// TIA Portal V20 export
DATA_BLOCK "OP2_DB"   // DB1
// stored: InstanceOfName OP2, InstanceOfType FB
"OP2"
   // VAR
   //    CONTROL_MAN : Struct
   //       B0 : Bool;
   //       B1 : Bool;
   //       B2 : Bool;
   //       B3 : Bool;
   //       B4 : Bool;
   //       B5 : Bool;
   //       B6 : Bool;
   //       B7 : Bool;
   //       B8 : Bool;
   //       B9 : Bool;
   //       odfuk_1 : Bool;
   //       odfuk_2 : Bool;
   //       B12 : Bool;
   //       B13 : Bool;
   //       B14 : Bool;
   //       B15 : Bool;
   //       B16 : Bool;
   //       B17 : Bool;
   //       B18 : Bool;
   //       B19 : Bool;
   //       B20 : Bool;
   //       B21 : Bool;
   //       B22 : Bool;
   //       B23 : Bool;
   //       B24 : Bool;
   //       B25 : Bool;
   //       B26 : Bool;
   //       B27 : Bool;
   //       B28 : Bool;
   //       B29 : Bool;
   //       B30 : Bool;
   //       B31 : Bool;
   //    END_STRUCT;
   //    CONTROL_AUTOMAT : Struct
   //       connect : Bool;
   //       send : Bool;
   //       reciv : Bool;
   //       trcv : Bool;
   //       discon : Bool;
   //       B5 : Bool;
   //       B6 : Bool;
   //       B7 : Bool;
   //       B8 : Bool;
   //       B9 : Bool;
   //       B10 : Bool;
   //       B11 : Bool;
   //       B12 : Bool;
   //       B13 : Bool;
   //       B14 : Bool;
   //       B15 : Bool;
   //       B16 : Bool;
   //       B17 : Bool;
   //       B18 : Bool;
   //       B19 : Bool;
   //       B20 : Bool;
   //       B21 : Bool;
   //       B22 : Bool;
   //       B23 : Bool;
   //       B24 : Bool;
   //       B25 : Bool;
   //       B26 : Bool;
   //       B27 : Bool;
   //       B28 : Bool;
   //       B29 : Bool;
   //       B30 : Bool;
   //       B31 : Bool;
   //    END_STRUCT;
   //    SENSORS : Struct
   //       S0 : Bool;
   //       S1 : Bool;
   //       S2 : Bool;
   //       S3 : Bool;
   //       S4 : Bool;
   //       S5 : Bool;
   //       S6 : Bool;
   //       S7 : Bool;
   //       S8 : Bool;
   //       S9 : Bool;
   //       S10 : Bool;
   //       S11 : Bool;
   //       S12 : Bool;
   //       S13 : Bool;
   //       S14 : Bool;
   //       S15 : Bool;
   //       S16 : Bool;
   //       S17 : Bool;
   //       S18 : Bool;
   //       S19 : Bool;
   //       S20 : Bool;
   //       S21 : Bool;
   //       S22 : Bool;
   //       S23 : Bool;
   //       S24 : Bool;
   //       S25 : Bool;
   //       S26 : Bool;
   //       S27 : Bool;
   //       S28 : Bool;
   //       S29 : Bool;
   //       S30 : Bool;
   //       S31 : Bool;
   //    END_STRUCT;
   //    SENSORS_1 : Struct
   //       S0 : Bool;
   //       S1 : Bool;
   //       S2 : Bool;
   //       S3 : Bool;
   //       S4 : Bool;
   //       S5 : Bool;
   //       S6 : Bool;
   //       S7 : Bool;
   //       S8 : Bool;
   //       S9 : Bool;
   //       S10 : Bool;
   //       S11 : Bool;
   //       S12 : Bool;
   //       S13 : Bool;
   //       S14 : Bool;
   //       S15 : Bool;
   //       S16 : Bool;
   //       S17 : Bool;
   //       S18 : Bool;
   //       S19 : Bool;
   //       S20 : Bool;
   //       S21 : Bool;
   //       S22 : Bool;
   //       S23 : Bool;
   //       S24 : Bool;
   //       S25 : Bool;
   //       S26 : Bool;
   //       S27 : Bool;
   //       S28 : Bool;
   //       S29 : Bool;
   //       S30 : Bool;
   //       S31 : Bool;
   //    END_STRUCT;
   //    S_0 : "SENSOR";
   //    S_1 : "SENSOR";
   //    S_2 { S7_SetPoint := 'True'} : "SENSOR";
   //    S_3 { S7_SetPoint := 'True'} : "SENSOR";
   //    S_4 { S7_SetPoint := 'True'} : "SENSOR";
   //    S_5 { S7_SetPoint := 'True'} : "SENSOR";
   //    S_6 { S7_SetPoint := 'True'} : "SENSOR";
   //    S_7 { S7_SetPoint := 'True'} : "SENSOR";
   //    S_8 { S7_SetPoint := 'True'} : "SENSOR";
   //    S_9 { S7_SetPoint := 'True'} : "SENSOR";
   //    S_10 { S7_SetPoint := 'True'} : "SENSOR";
   //    S_11 { S7_SetPoint := 'True'} : "SENSOR";
   //    S_12 { S7_SetPoint := 'True'} : "SENSOR";
   //    S_13 { S7_SetPoint := 'True'} : "SENSOR";
   //    S_14 { S7_SetPoint := 'True'} : "SENSOR";
   //    S_15 { S7_SetPoint := 'True'} : "SENSOR";
   //    S_16 { S7_SetPoint := 'True'} : "SENSOR";
   //    M_1 : "MOTOR_CONTROL_BLOCK";
   //    M_2 { S7_SetPoint := 'True'} : "MOTOR_CONTROL_BLOCK";
   //    M_3 { S7_SetPoint := 'True'} : "MOTOR_CONTROL_BLOCK";
   //    SQCR { S7_SetPoint := 'True'} : Int;
   //    hmi_sqcr : Int;
   //    TRIG : Struct
   //       inicial_ok_op : Bool;
   //       T2 : Bool;
   //       T3 : Bool;
   //       T4 : Bool;
   //       T5 : Bool;
   //       T6 : Bool;
   //       T7 : Bool;
   //       T8 : Bool;
   //       T9 : Bool;
   //       T10 : Bool;
   //       T11 : Bool;
   //       T12 : Bool;
   //       T13 : Bool;
   //       T14 : Bool;
   //       T15 : Bool;
   //       T16 : Bool;
   //       op_1_ready : Bool;
   //    END_STRUCT;
   //    MEMOR : Struct
   //       n_trig_vypnuti : Bool;
   //       M1 : Bool;
   //       M2 : Bool;
   //       M3 : Bool;
   //       M4 : Bool;
   //       p_trig_odavacka : Bool;
   //       M6 : Bool;
   //       M7 : Bool;
   //       M8 : Bool;
   //       M9 : Bool;
   //       M10 : Bool;
   //       M11 : Bool;
   //       RESET_ERROR : Bool;
   //       M13 : Bool;
   //       M14 : Bool;
   //       M15 : Bool;
   //       SETOVANI_START : Bool;
   //       M17 : Bool;
   //       M18 : Bool;
   //       M19 : Bool;
   //       M20 : Bool;
   //       M21 : Bool;
   //       M22 : Bool;
   //       M23 : Bool;
   //       M24 : Bool;
   //       M25 : Bool;
   //       M26 : Bool;
   //       M27 : Bool;
   //       M28 : Bool;
   //       M29 : Bool;
   //       M30 : Bool;
   //       N_TRIG_SAFETY : Bool;
   //       M32 : Bool;
   //       M33 : Bool;
   //       start_caklu : Bool;
   //       M35 : Bool;
   //       M36 : Bool;
   //       M37 : Bool;
   //       M38 : Bool;
   //       M39 : Bool;
   //       ALARM_GLOBAL : Bool;
   //       M41 : Bool;
   //       M42 : Bool;
   //       M43 : Bool;
   //       M44 : Bool;
   //       M45 : Bool;
   //       M46 : Bool;
   //       M47 : Bool;
   //       M48 : Bool;
   //       M49 : Bool;
   //       wrong_p_trig : Bool;
   //       alarm_p_trig : Bool;
   //       M52 : Bool;
   //       M53 : Bool;
   //       M54 : Bool;
   //       M55 : Bool;
   //       M56 : Bool;
   //       M57 : Bool;
   //       M58 : Bool;
   //       M59 : Bool;
   //       M60 : Bool;
   //       M61 : Bool;
   //       M62 : Bool;
   //       M63 : Bool;
   //    END_STRUCT;
   //    "TIMER" : Struct
   //       TIMER_0 : IEC_TIMER;
   //       TIMER_1 : IEC_TIMER;
   //       TIMER_2 : IEC_TIMER;
   //       TIMER_3 : IEC_TIMER;
   //       TIMER_4 : IEC_TIMER;
   //       air : IEC_TIMER;
   //       TIMER_6 : IEC_TIMER;
   //       TIMER_7 : IEC_TIMER;
   //    END_STRUCT;
   //    HMI : Struct
   //       povoleni_volby_receptu : Bool;
   //       "svetlo_on/off" : Bool;
   //       ALARM_VIDITELNOST : Bool;
   //       hmi_3 : Bool;
   //       hmi_4 : Bool;
   //       hmi_5 : Bool;
   //       hmi_6 : Bool;
   //       hmi_7 : Bool;
   //       hmi_8 : Bool;
   //       hmi_9 : Bool;
   //       hmi_10 : Bool;
   //       hmi_11 : Bool;
   //       hmi_12 : Bool;
   //       hmi_13 : Bool;
   //       hmi_14 : Bool;
   //       hmi_15 : Bool;
   //    END_STRUCT;
   //    int_hodnota_zpravy { ExternalAccessible := 'False'; ExternalVisible := 'False'; ExternalWritable := 'False'} : Word;
   //    CTRV_LEN { ExternalAccessible := 'False'; ExternalVisible := 'False'; ExternalWritable := 'False'} : UDInt;
   //    TCON_Instance { S7_SetPoint := 'True'} : TCON;
   //    TSEND_Instance { S7_SetPoint := 'True'} : TSEND;
   //    TRCV_Instance { S7_SetPoint := 'True'} : TRCV;
   //    TDISCON_Instance { S7_SetPoint := 'True'} : TDISCON;
   //    Tisk : Struct
   //       pole2_index_bajt : Int := 14;
   //       pole2_index_hodnota : Byte := 16#02;
   //       datum_chyba : Bool;
   //       pole2_kratky : Bool;
   //       jeden_ramec : Bool := true;
   //    END_STRUCT;
   // END_VAR
BEGIN
END_DATA_BLOCK
